{attribute 'linkalways'} 
{attribute 'no_explicit_call' := 'This FB is a CLASS and must be accessed using methods or properties'}
{attribute 'enable_dynamic_creation'}
FUNCTION_BLOCK _Array0to2OfTcVnPoint2_REAL EXTENDS ArrayDatatypeBase_1D
VAR CONSTANT
	lBound : DINT := 0;
	uBound : DINT := 2;
END_VAR
VAR
	localData : ARRAY [lBound..uBound] OF TcVnPoint2_REAL;
	activeData : REFERENCE TO ARRAY [lBound..uBound] OF TcVnPoint2_REAL REF= localData;
	elements : ARRAY [lBound..uBound] OF _TcVnPoint2_REAL;
	baseType : _TcVnPoint2_REAL;
END_VAR

PROPERTY PUBLIC Address : PVOID
GET
Address := ADR(activeData);
END_GET
END_PROPERTY

PROPERTY PUBLIC BaseDatatype : I_Datatype
GET
BaseDatatype := baseType;
END_GET
END_PROPERTY

METHOD PUBLIC ClearReference
VAR_INPUT
END_VAR
activeData REF= localData;
SetElementReference();
END_METHOD

METHOD PUBLIC Clone : I_Datatype
VAR
    pClone : POINTER TO _Array0to2OfTcVnPoint2_REAL;
END_VAR
pClone := __NEW(_Array0to2OfTcVnPoint2_REAL());
pClone^.Value := Value;
Clone := pClone^;
END_METHOD

METHOD FB_init : BOOL
VAR_INPUT
	bInitRetains : BOOL; // if TRUE, the retain variables are initialized (warm start / cold start)
	bInCopyCode : BOOL;  // if TRUE, the instance afterwards gets moved into the copy code (online change)
END_VAR
SetElementReference();
END_METHOD

METHOD PUBLIC MakeReferenceTo
VAR_INPUT
	ReferenceTarget : REFERENCE TO ARRAY [lBound..uBound] OF TcVnPoint2_REAL;
END_VAR
activeData REF= ReferenceTarget;
SetElementReference();
END_METHOD

METHOD PROTECTED OnSerializeArrayValues
VAR_INPUT
	Serializer : I_Serializer;
END_VAR
VAR
	i : DINT;
END_VAR
FOR i := lBound TO uBound DO
	elements[i].SerializeWith(Serializer);
END_FOR
END_METHOD

METHOD PROTECTED SetElementReference
VAR_INPUT
END_VAR
VAR
	i : DINT;
END_VAR
FOR i := lBound TO uBound DO
	elements[i].MakeReferenceTo(activeData[i]);
END_FOR
END_METHOD

PROPERTY PUBLIC Size : UDINT
GET
Size := SIZEOF(activeData);
END_GET
END_PROPERTY

METHOD PROTECTED TryDeserializeArrayValues : BOOL
VAR_INPUT
	Deserializer : I_Deserializer;
	Feedback : I_DeserializerFeedback;
END_VAR
VAR
	failed : BOOL;
	enumerator : I_DeserializerArrayForwardEnumerator;
	i : DINT;
END_VAR
enumerator := Deserializer.GetArrayEnumerator();
i := lBound;

WHILE enumerator.MoveNext() AND i <= uBound AND NOT failed DO
	
	IF NOT elements[i].TryDeserializeFrom(enumerator.Current, Feedback) THEN
		failed := TRUE;
		EXIT;
	END_IF
	i := i + 1;

END_WHILE
enumerator.Dispose();

TryDeserializeArrayValues := NOT failed;
END_METHOD

METHOD PUBLIC TryGetElementAsDatatypeByIndex : BOOL
VAR_INPUT
	Index : DINT;
	Destination : REFERENCE TO I_Datatype;
END_VAR
IF Index < lbound OR Index > ubound THEN
	RETURN;
END_IF

Destination := elements[Index];
TryGetElementAsDatatypeByIndex := TRUE;
END_METHOD

METHOD PUBLIC TryGetLowerBound : BOOL
VAR_INPUT
	Dimention : UDINT;
	Destination : REFERENCE TO DINT;
END_VAR
IF Dimention = 1 THEN
	Destination := lBound;
	TryGetLowerBound := TRUE;
END_IF
END_METHOD

METHOD PUBLIC TryGetUpperBound : BOOL
VAR_INPUT
	Dimention : UDINT;
	Destination : REFERENCE TO DINT;
END_VAR
IF Dimention = 1 THEN
	Destination := uBound;
	TryGetUpperBound := TRUE;
END_IF
END_METHOD

METHOD TryMakeReferenceTo : BOOL
VAR_INPUT
	Target : I_Datatype;
END_VAR
VAR
	pTargetData : POINTER TO ARRAY [lBound..uBound] OF TcVnPoint2_REAL;
END_VAR
IF NOT IsEquivalentTo(Target) THEN
	RETURN;
END_IF

pTargetData := Target.Address;
activeData REF= pTargetData^;
SetElementReference();
TryMakeReferenceTo := TRUE;
END_METHOD

PROPERTY PUBLIC Value : REFERENCE TO ARRAY [lBound..uBound] OF TcVnPoint2_REAL;
GET
Value ref= activeData;
END_GET
END_PROPERTY

END_FUNCTION_BLOCK

(* stored: Version 1.1.0.1, ProductVersion 3.1.4024.13
   POU _Array0to2OfTcVnPoint2_REAL: Id {95a1f11c-7b3e-0adb-266b-051ed318cba3}, SpecialFunc None
   Folder Core: Id {b5607c07-a63f-05a1-0d9a-7af94a562e8a}
   Folder Constructor: Id {934e84b2-ce2f-0590-3406-126821dce628}
   Folder Protected: Id {6dd3ecbd-0c29-0d84-2b84-f774249a5cd9}
   Folder Customize: Id {778cb6b6-8384-0a2c-20bc-2f52a7e87782}
   Property Address: Id {2e7ec9bd-62c5-0735-0f45-b6855f9c5272}
   Get Get: Id {a75ea913-9b91-046f-3a53-b92f59742d11}
   Property BaseDatatype: Id {1d7ee3a8-9932-0cab-368a-d07f5ffae6e8}
   Get Get: Id {5f514769-7984-051c-24a6-abc7d2cc7c05}
   Method ClearReference: Id {3e623531-6c7e-0504-36bb-90a6f3a09482}
   Method Clone: Id {fee38ac9-62cb-012d-292c-18cc4da335ca}
   Method FB_init: Id {8b52167d-9a03-07c9-0a33-8cc3916ea438}
   Method MakeReferenceTo: Id {9388318d-513a-0449-1d0f-2e39a830ce48}
   Method OnSerializeArrayValues: Id {62646663-497d-0ba1-065b-5e9f71f991d3}
   Method SetElementReference: Id {9e447a9b-10f1-0ad1-3558-523ee4739146}
   Property Size: Id {4f73b033-68ca-0bc1-01a1-d3fe5db2756e}
   Get Get: Id {f589a200-a8f6-0a4b-1b40-3e9697210a9f}
   Method TryDeserializeArrayValues: Id {82a3dfe3-0622-0b67-2f5d-04d5d880d118}
   Method TryGetElementAsDatatypeByIndex: Id {77fda498-8b87-02fb-0ceb-6dc63d44c08f}
   Method TryGetLowerBound: Id {c8118e29-7b67-028d-2264-1426eef1915d}
   Method TryGetUpperBound: Id {bdd2a971-de8f-0931-27d7-c6e61414fb68}
   Method TryMakeReferenceTo: Id {f7101726-5a76-049b-2c83-0ca4951f2a8e}
   Property Value: Id {21c30b35-d46a-0f72-2dff-e254c19a71fa}
   Get Get: Id {3500656b-d5d4-018e-154e-35bce26832ac} *)
